FUNCTION_BLOCK BasicTest (* Basic FB with an ECC *)
  (* Standard: 61499-1; Classification: Fixture; ApplicationDomain: Testing; Function: Exercise import/export; Type: Basic FB; Description: Copyright (c) 2026 Martin Erich Jobst This program and the accompanying materials are made available under the terms of the Eclipse Public License 2.0 which is available at https://www.eclipse.org/legal/epl-2.0/ SPDX-License-Identifier: EPL-2.0 *)
  (* Version 1.0, 2026-10-23, Martin Jobst, Eclipse, Canonical fixture *)
  PACKAGE fixture::basic;
  IMPORT fixture;
  (* Compiler header: basic.h *)
  (* Compiler classdef: BasicTest *)
  (* Compiler C Eclipse 4diac 1.0 *)
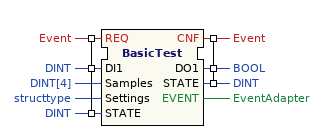
  EVENT_INPUT
    REQ WITH DI1, STATE; (* Request *)
  END_EVENT
  EVENT_OUTPUT
    CNF WITH DO1, STATE; (* Confirmation *)
  END_EVENT
  VAR_INPUT
    DI1 : DINT := DINT#1; {SET_ATTRIBUTE(IntegerAttribute, 1)} {SET_ATTRIBUTE(StructuredAttribute, (7,TRUE,'fixture'))}
    Samples : ARRAY [0..3] OF DINT;
    Settings : structtype;
  END_VAR
  VAR_OUTPUT
    DO1 : BOOL;
  END_VAR
  VAR_IN_OUT
    STATE : DINT := DINT#0;
  END_VAR
  PLUGS
    EVENT : EventAdapter(REQD := WSTRING#'request'); (* Event/data adapter *) {SET_ATTRIBUTE(AdapterAttribute, AdapterValue)}
  END_PLUGS
  VAR CONSTANT
    limit : DINT := DINT#10;
  END_VAR
  VAR
    counter : DINT := DINT#0;
  END_VAR
  FBS
    helper : SimpleTest; (* Internal helper *)
  END_FBS
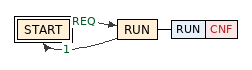
  EC_STATES
    START; (* Initial State *)
    RUN : RUN -> CNF;
  END_STATES
  EC_TRANSITIONS
    START TO RUN := REQ;
    RUN TO START := 1;
  END_TRANSITIONS
  ALGORITHM RUN IN ST:
	DO1 := DI1 > 0;
  END_ALGORITHM
  ALGORITHM SCRIPT IN Lua:
emit("fixture")
  END_ALGORITHM
  METHOD Compute : DINT (* Computes a value *)
  VAR_INPUT
    operand : DINT;
  END_VAR
  VAR_OUTPUT
    offset : DINT;
  END_VAR
Compute := operand + offset;
  END_METHOD
  METHOD ScriptMethod : DINT
  VAR_INPUT
    operand : DINT;
  END_VAR
  VAR_OUTPUT
    result : DINT;
  END_VAR
return operand
  END_METHOD
END_FUNCTION_BLOCK
